{region 'Documentation'}
(*!
<summary>Checks that at least one selected bit is FALSE.</summary>
*)
{endregion}
FUNCTION_BLOCK AssertContainsFalse_LWord EXTENDS AssertionBase
VAR_INPUT
    IN : LWORD; //! Actual bitfield.
    Mask : LWORD := 16#FFFFFFFFFFFFFFFF; //! Selects evaluated bits; defaults to all bits. An empty mask produces Error during evaluation.
END_VAR

SUPER^();

{region 'Documentation'}
(*!
<summary>Rejects an empty mask before checking for a matching selected bit.</summary>
*)
{endregion}
METHOD PROTECTED Assert
VAR
    Message : STRING(GVL_Constants.MessageLength);
    MaskText : STRING(GVL_Constants.AssertionValueLength);
    ActualText : STRING(GVL_Constants.AssertionValueLength);
END_VAR
VAR CONSTANT
    NoMask : LWORD := 16#00;
    HexDigitCount : USINT := 16;
END_VAR
IF NOT EvaluationActive THEN
    RETURN;
END_IF;

IF Result = E_Result.Error THEN
    RETURN;
END_IF;

IF Mask = NoMask THEN
    MaskText := CreateAssertionTextValue_Hex(Value := Mask,
        DigitCount := HexDigitCount);
    Message := CONCAT('Assertion error: mask must not be empty. Mask = ',
        MaskText);
    Message := CONCAT(Message, '.');
    Error(Message := Message);
    RETURN;
END_IF;

IF Result = E_Result.Failed THEN
    RETURN;
END_IF;

IF (IN AND Mask) = Mask THEN
    MaskText := CreateAssertionTextValue_Hex(Value := Mask,
        DigitCount := HexDigitCount);
    ActualText := CreateAssertionTextValue_Hex(Value := IN,
        DigitCount := HexDigitCount);
    Message := CONCAT('Assertion failed: no selected bit is FALSE. Mask = ',
        MaskText);
    Message := CONCAT(Message, ', Actual = ');
    Message := CONCAT(Message, ActualText);
    Message := CONCAT(Message, '.');
    Fail(Message := Message);
    RETURN;
END_IF;

Pass();
END_METHOD

END_FUNCTION_BLOCK

(* stored: Version 1.1.0.1
   POU AssertContainsFalse_LWord: Id {9682cfef-f958-48c9-8686-aebf0a5665d3}, SpecialFunc None
   Folder Internal: Id {cd91c6af-4591-4d7f-a887-def12718b77e}
   Method Assert: Id {12fa3551-d541-4812-a2c6-757da7698f6f} *)
